Fanuc KAREL source: KT00477.KL

PROGRAM KT00477
%NOLOCKGROUP
VAR
  P1: POSITION
  P2: POSITION
  OUT: JOINTPOS
BEGIN
  OUT = P1 : P2
END KT00477
